(* IEC 61131-3 sources: Elmo_Master/Lasal_PRG/Welcon8Axis_EtherCAT_Test_With_RobotAxis/Network/DS402_Network, 1 file *)

(* ---- ONE_DS402_Network_Table.st ---- *)
#define OBJECTS_CONFIG

//Define part of class DriveAxisDS402
//=============================================================================================
//Timeouts / Thresholds
//=============================================================================================
#define ECAT_DRIVE_ENABLE_TIMEOUT 1000

FUNCTION GLOBAL TAB ONE_DS402_Network
-1$UINT, 0$UINT,
0$UINT, 0$UINT,

2$UDINT,
TO_UDINT(4054914251), "DriveAxisDS402", 1$UINT, 3$UINT, 4$UINT,
TO_UDINT(595672599), "DriveAxisDS402_Base", 1$UINT, 0$UINT, 0$UINT,

_NO_ATTR, TO_UDINT(4273818432), "DRIVEAXISDS402_AXIS2",
_NO_ATTR, TO_UDINT(400486005), "DRIVEAXISDS402_AXIS4",
_NO_ATTR, TO_UDINT(4191194969), "DRIVEAXISDS402_AXIS6",
_NO_ATTR, TO_UDINT(510173790), "DRIVEAXISDS402_AXIS8",

//Internal connections
0$UDINT,
0$UDINT,
0$UDINT,
0$UDINT,

//Initialization values
0$UDINT,
4$UDINT,
TO_UDINT(0), "SetOpMode", TO_UDINT(8),//|DS402_Network.DriveAxisDS402_Axis2.SetOpMode;
TO_UDINT(1), "SetOpMode", TO_UDINT(8),//|DS402_Network.DriveAxisDS402_Axis4.SetOpMode;
TO_UDINT(2), "SetOpMode", TO_UDINT(8),//|DS402_Network.DriveAxisDS402_Axis6.SetOpMode;
TO_UDINT(3), "SetOpMode", TO_UDINT(8),//|DS402_Network.DriveAxisDS402_Axis8.SetOpMode;

//Symbolic initialization values
0$UDINT,
0$UDINT,

//Initialization of string values
0$UDINT,
0$UDINT,

//Configuration of tasks (RealTime, Cyclic, Background)
0$UDINT,
4$UDINT,
TO_UDINT(0), (1)$UDINT, 4194303$DINT, 	//DRIVEAXISDS402_AXIS2
TO_UDINT(1), (1)$UDINT, 4194303$DINT, 	//DRIVEAXISDS402_AXIS4
TO_UDINT(2), (1)$UDINT, 4194303$DINT, 	//DRIVEAXISDS402_AXIS6
TO_UDINT(3), (1)$UDINT, 4194303$DINT, 	//DRIVEAXISDS402_AXIS8

0$UDINT,
0$UDINT,

0$UDINT,
0$UDINT,

//External connections
0$UDINT,
44$UDINT,
TO_UDINT(0), "CiA_ControlWord", C_DIR, TO_UDINT(3391823300), "WELCON_11","RxPDO9_Controlword2",
TO_UDINT(0), "CiA_StatusWord", C_DIR, TO_UDINT(3391823300), "WELCON_11","TxPDO9_Statusword2",
TO_UDINT(0), "ModesOfOperation", C_TRY, TO_UDINT(3391823300), "WELCON_11","RxPDO9_ModesOfOperation2",
TO_UDINT(0), "ModesOfOperationDisplay", C_TRY, TO_UDINT(3391823300), "WELCON_11","TxPDO9_ModesOfOperationDisplay2",
TO_UDINT(0), "PositionActualValue", C_TRY, TO_UDINT(3391823300), "WELCON_11","TxPDO9_PositionActualValue2",
TO_UDINT(0), "TargetPosition", C_TRY, TO_UDINT(3391823300), "WELCON_11","RxPDO9_TargetPosition2",
TO_UDINT(0), "TargetTorque", C_TRY, TO_UDINT(3391823300), "WELCON_11","RxPDO9_TargetTorque2",
TO_UDINT(0), "TargetVelocity", C_TRY, TO_UDINT(3391823300), "WELCON_11","RxPDO9_TargetVelocity2",
TO_UDINT(0), "TorqueActualValue", C_TRY, TO_UDINT(3391823300), "WELCON_11","TxPDO9_TorqueActualValue2",
TO_UDINT(0), "VelocityActualValue", C_TRY, TO_UDINT(3391823300), "WELCON_11","TxPDO9_VelocityActualValue2",
TO_UDINT(0), "Online", C_TRY, TO_UDINT(3391823300), "WELCON_11","Online",
TO_UDINT(1), "CiA_ControlWord", C_DIR, TO_UDINT(3775286791), "WELCON_21","RxPDO9_Controlword2",
TO_UDINT(1), "CiA_StatusWord", C_DIR, TO_UDINT(3775286791), "WELCON_21","TxPDO9_Statusword2",
TO_UDINT(1), "ModesOfOperation", C_TRY, TO_UDINT(3775286791), "WELCON_21","RxPDO9_ModesOfOperation2",
TO_UDINT(1), "ModesOfOperationDisplay", C_TRY, TO_UDINT(3775286791), "WELCON_21","TxPDO9_ModesOfOperationDisplay2",
TO_UDINT(1), "PositionActualValue", C_TRY, TO_UDINT(3775286791), "WELCON_21","TxPDO9_PositionActualValue2",
TO_UDINT(1), "TargetPosition", C_TRY, TO_UDINT(3775286791), "WELCON_21","RxPDO9_TargetPosition2",
TO_UDINT(1), "TargetTorque", C_TRY, TO_UDINT(3775286791), "WELCON_21","RxPDO9_TargetTorque2",
TO_UDINT(1), "TargetVelocity", C_TRY, TO_UDINT(3775286791), "WELCON_21","RxPDO9_TargetVelocity2",
TO_UDINT(1), "TorqueActualValue", C_TRY, TO_UDINT(3775286791), "WELCON_21","TxPDO9_TorqueActualValue2",
TO_UDINT(1), "VelocityActualValue", C_TRY, TO_UDINT(3775286791), "WELCON_21","TxPDO9_VelocityActualValue2",
TO_UDINT(1), "Online", C_TRY, TO_UDINT(3775286791), "WELCON_21","Online",
TO_UDINT(2), "CiA_ControlWord", C_DIR, TO_UDINT(4162682694), "WELCON_31","RxPDO9_Controlword2",
TO_UDINT(2), "CiA_StatusWord", C_DIR, TO_UDINT(4162682694), "WELCON_31","TxPDO9_Statusword2",
TO_UDINT(2), "ModesOfOperation", C_TRY, TO_UDINT(4162682694), "WELCON_31","RxPDO9_ModesOfOperation2",
TO_UDINT(2), "ModesOfOperationDisplay", C_TRY, TO_UDINT(4162682694), "WELCON_31","TxPDO9_ModesOfOperationDisplay2",
TO_UDINT(2), "PositionActualValue", C_TRY, TO_UDINT(4162682694), "WELCON_31","TxPDO9_PositionActualValue2",
TO_UDINT(2), "TargetPosition", C_TRY, TO_UDINT(4162682694), "WELCON_31","RxPDO9_TargetPosition2",
TO_UDINT(2), "TargetTorque", C_TRY, TO_UDINT(4162682694), "WELCON_31","RxPDO9_TargetTorque2",
TO_UDINT(2), "TargetVelocity", C_TRY, TO_UDINT(4162682694), "WELCON_31","RxPDO9_TargetVelocity2",
TO_UDINT(2), "TorqueActualValue", C_TRY, TO_UDINT(4162682694), "WELCON_31","TxPDO9_TorqueActualValue2",
TO_UDINT(2), "VelocityActualValue", C_TRY, TO_UDINT(4162682694), "WELCON_31","TxPDO9_VelocityActualValue2",
TO_UDINT(2), "Online", C_TRY, TO_UDINT(4162682694), "WELCON_31","Online",
TO_UDINT(3), "CiA_ControlWord", C_DIR, TO_UDINT(3076319617), "WELCON_41","RxPDO9_Controlword2",
TO_UDINT(3), "CiA_StatusWord", C_DIR, TO_UDINT(3076319617), "WELCON_41","TxPDO9_Statusword2",
TO_UDINT(3), "ModesOfOperation", C_TRY, TO_UDINT(3076319617), "WELCON_41","RxPDO9_ModesOfOperation2",
TO_UDINT(3), "ModesOfOperationDisplay", C_TRY, TO_UDINT(3076319617), "WELCON_41","TxPDO9_ModesOfOperationDisplay2",
TO_UDINT(3), "PositionActualValue", C_TRY, TO_UDINT(3076319617), "WELCON_41","TxPDO9_PositionActualValue2",
TO_UDINT(3), "TargetPosition", C_TRY, TO_UDINT(3076319617), "WELCON_41","RxPDO9_TargetPosition2",
TO_UDINT(3), "TargetTorque", C_TRY, TO_UDINT(3076319617), "WELCON_41","RxPDO9_TargetTorque2",
TO_UDINT(3), "TargetVelocity", C_TRY, TO_UDINT(3076319617), "WELCON_41","RxPDO9_TargetVelocity2",
TO_UDINT(3), "TorqueActualValue", C_TRY, TO_UDINT(3076319617), "WELCON_41","TxPDO9_TorqueActualValue2",
TO_UDINT(3), "VelocityActualValue", C_TRY, TO_UDINT(3076319617), "WELCON_41","TxPDO9_VelocityActualValue2",
TO_UDINT(3), "Online", C_TRY, TO_UDINT(3076319617), "WELCON_41","Online",

//Magic internal connections
0$UDINT,
0$UDINT,

//Configuration of timeslots of tasks (RealTime, Cyclic)
#ifdef __LSLLDR_TIMESLOTS__
0$UDINT,
0$UDINT,

0$UDINT,
0$UDINT,

#endif //__LSLLDR_TIMESLOTS__

//MultiMaster connections
#ifdef __LSLLDR_MULTIMASTER__
0$UDINT,
0$UDINT,
#endif //__LSLLDR_MULTIMASTER__

//Configuration for task ID (RealTime, CyclicTime)
#ifdef __LSLLDR_TASKID__
"\\\\TASKS2  "
0$UDINT,
4$UDINT,
(0)$UDINT, 	//DRIVEAXISDS402_AXIS2
(0)$UDINT, 	//DRIVEAXISDS402_AXIS4
(0)$UDINT, 	//DRIVEAXISDS402_AXIS6
(0)$UDINT, 	//DRIVEAXISDS402_AXIS8

0$UDINT,
0$UDINT,

0$UDINT,
0$UDINT,

#endif //__LSLLDR_TASKID__

END_FUNCTION
